{attribute 'qualified_only'}
VAR_GLOBAL
	//ST_TwinSAFE_IN
	stTwinSAFE_OUT	AT %Q* :ST_TwinSAFE_OUT;
	stTwinSAFE_IN	AT %I* : ST_TwinSAFE_IN;
	DoorMonitorFromPLC AT %I* : BOOL;
	SolonoidStatus AT %I* : BOOL;
END_VAR

(* stored: Version 1.1.0.1, ProductVersion 3.1.4026.18
   GVL GVL_Safety: Id {0521510e-a6b2-4216-9dd3-0a59704f168a} *)
